(* PLC project DemoProject, Voltrus Voltrus Studio 1.0 *)
(* stored: creationDateTime 2026-09-13T00:00:00 *)

TYPE Recipe : STRUCT
  target : REAL;
  enabled : BOOL;
  label : STRING(16);
END_STRUCT;
END_TYPE

TYPE SpeedLimit : INT(0..100);
END_TYPE

PROGRAM Main
  VAR_INPUT
    start_cmd : BOOL := FALSE;
  END_VAR
  VAR_OUTPUT
    running : BOOL;
  END_VAR
  VAR_IN_OUT
    recipe : Recipe;
  END_VAR
  VAR
    cycle_count : DINT := 0;
    delay : TON;
  END_VAR

            
running := start_cmd;
cycle_count := cycle_count + 1;
recipe.target := recipe.target * 2.0;
delay(IN := start_cmd, PT := T#10MS);
            
          
END_PROGRAM

CONFIGURATION Config0
  RESOURCE Res0 ON PLC
    TASK MainTask(INTERVAL := T#20ms, PRIORITY := 0);
    PROGRAM Main_Instance WITH MainTask : Main;
  END_RESOURCE
END_CONFIGURATION
